Fanuc KAREL source: kd00007.KL

-- PROVISIONAL review KL for V770-1; original PC SHA256 c8d788d161ffa7bbdaee540d95ec0536ce15f6d7225dbdac346538f178e11269
-- Incomplete behavior may be omitted. Consult companion uncertainty JSON. Do not deploy.
PROGRAM KD00007
%NOLOCKGROUP
-- UNRESOLVED_DECL I type=020010
-- UNRESOLVED_DECL J type=020010
-- UNRESOLVED_DECL B type=020012
-- UNRESOLVED_DECL R type=020011
-- UNRESOLVED_DECL S type=021f50
BEGIN
  -- UNRESOLVED_PC offsets 5-12; opcodes 9D,23
  -- UNRESOLVED_PC offsets 17-21; opcodes 7F
END KD00007
